Universal Robots URScript: swab_sampling.script

global swab_poses=make_list(0,0,6)
global pose_list_hor=make_list(0,0,420)
global pose_list_ver=make_list(0,0,420)
global cntd=False
global trgt_waypts=make_list(0,0,6)
global new_z=0
global first_pts=make_list(0,0,15)
global temp_pose_force=p[0,0,0,0,0,0]
global delta_rx=0
global new_dz=0
global server_msg=""
global delta_x=0
global delta_y=0


def connect2server():
	IP="192.168.12.139"
	port=3002
	while(cntd==False):
		cntd=socket_open(IP,port)
		if(cntd==True):
			textmsg("Connected to server")
		end
	end
	socket_send_string("SCAN_TARGET")
end


def get_hor_pose_from_server():

	IP="192.168.12.139"
	port=3002
	if(cntd==True):
		textmsg("Connected to server")
	end
	while(cntd==False):
		cntd=socket_open(IP,port)
		if(cntd==True):
			textmsg("Connected to server")
		end
		sleep(0.2)
	end
	socket_send_string("GET_POSE_HOR")
	idx=socket_read_ascii_float(1,timeout=-1)
	textmsg("Index from server=",idx[1])
	itn_i=0
	while(itn_i<idx[1]):
		msg=socket_read_ascii_float(6,timeout=-1)
		i=1
		while(i<7):
			swab_poses.append(msg[i])
			i=i+1
		end
		pose_list_hor.extend(swab_poses)
		swab_poses.clear()
		socket_send_string("OK")
		itn_i=itn_i+1
	end
	socket_read_line(timeout=-1)
	if(cntd==True):
		cntd=False
		socket_close()
	end
	#textmsg("server msg",swab_poses)
	textmsg("pose list",pose_list_hor)
end


def get_ver_pose_from_server():
	IP="192.168.12.139"
	port=3002
	if(cntd==True):
		textmsg("Connected to server")
	end
	while(cntd==False):
		cntd=socket_open(IP,port)
		if(cntd==True):
			textmsg("Connected to server")
		end
		sleep(0.2)
	end
	socket_send_string("GET_POSE_VER")
	idx=socket_read_ascii_float(1,timeout=-1)
	textmsg("Index from server=",idx[1])
	itn_i=0
	while(itn_i<idx[1]):
		msg=socket_read_ascii_float(6,timeout=-1)
		i=1
		while(i<7):
			swab_poses.append(msg[i])
			i=i+1
		end
		pose_list_ver.extend(swab_poses)
		swab_poses.clear()
		socket_send_string("OK")
		itn_i=itn_i+1
	end
	socket_read_line(timeout=-1)
	if(cntd==True):
		cntd=False
		socket_close()
	end
	#textmsg("server msg",swab_poses)
	textmsg("pose list",pose_list_ver)
end


def move_to_first_point(code):
	first_pts.clear()
	k=0
	i=1
	l=1
	blend_r=0
	while(i<3):
		j=1
		while(j<=6):
			k=l-1
			if(code==1):
				first_pts.append(pose_list_hor[k])
			elif(code==2):
				first_pts.append(pose_list_ver[k])
			end
			j=j+1
			l=l+1
		end
		i=i+1
	end
	movel(p[first_pts[0]-delta_y,first_pts[1]+delta_x,first_pts[2],first_pts[3],first_pts[4],first_pts[5]],a=0.5,v=0.05,r=blend_r)
	sleep(2)
	zero_ftsensor()
	sleep(2)
	tcp_f=get_tcp_force()
	textmsg("Force after zeroing:",tcp_f)
	ftmode=True
	while(ftmode==True):
		tcp_f=get_tcp_force()
		if tcp_f[2]<0.7:
			speedl([0,0,-0.001,0,0,0],0.05,t=0.5)
		else:
			stopl(3)
			new_p=get_actual_tcp_pose()
			new_z=new_p[2]-first_pts[2]
			ftmode=False
		end
		sleep(0.2)
	end
	movel(p[first_pts[6]-delta_y,first_pts[7]+delta_x,first_pts[8]+new_z,first_pts[9],first_pts[10],first_pts[11]],a=0.5,v=0.05,r=blend_r)
	curr_tcp=get_actual_tcp_pose()
	textmsg("Current TCP",curr_tcp)
	#tcp_str=to_string(curr_tcp)
	popup("Tcp change",blocking=True)
	#temp_pose_force=p[first_pts[0],first_pts[1],first_pts[2],first_pts[3],first_pts[4],first_pts[5]]
	temp_pt=first_pts[2]
	first_pts.clear()
	zero_ftsensor()
	sleep(2)
	tcp_f=get_tcp_force()
	textmsg("Force after zeroing:",tcp_f)
	ftmode=True
	#ftmode=False
	while(ftmode==True):
		tcp_f=get_tcp_force()
		textmsg("Force",tcp_f)
		if tcp_f[2]<2.5:
			speedl([0,0,-0.005,0,0,0],0.05,t=0.5)
		else:
			stopl(3)
			new_p=get_actual_tcp_pose()
			new_dz=new_p[2]-temp_pt
			ftmode=False
			textmsg("DZ=",new_dz)
		end
		sleep(0.2)
	end
	IP="192.168.12.139"
	port=3002
	if(cntd==True):
		textmsg("Connected to server")
	end
	while(cntd==False):
		cntd=socket_open(IP,port)
		if(cntd==True):
			textmsg("Connected to server")
		end
		sleep(0.2)
	end
	socket_send_string("POSE")
	socket_send_string(str_cat("",curr_tcp))
	if(cntd==True):
		cntd=False
		socket_close()
	end

end

def follow_swab_trajectory_hor():
	idx=pose_list_hor.length()
	textmsg("idx",idx)
	idx=idx/6
	k=0
	i=3
	l=13
	delta_z=0.035
	zero_ftsensor()
	sleep(1)
	#tcp_f=get_tcp_force()
	#textmsg("Force at tip:",tcp_f)
	force_mode(temp_pose_force,[0,0,1,0,0,0],[0,0,0.3,0,0,0],2,[0.005,0.005,0.05,0.01,0.01,0.01])
	while(i<=idx):
		j=1
		while(j<=6):
			k=l-1
			trgt_waypts.append(pose_list_hor[k])
			j=j+1
			l=l+1
		end
		if(i<3):
			delta_rx=0
			delta_z=0
			blend_r=0
		elif((i-1)%5==0):
			blend_r=0
			delta_z=0.043
			#delta_rx=0.104
			delta_rx=0.3
		else:
			blend_r=0.002
			delta_z=0.043
			#delta_rx=0.104
			delta_rx=0.3
		end
		if(i==1):
			delta_z=0.005
			trgt_waypts[2]=trgt_waypts[2]+delta_z
		movel(p[trgt_waypts[0],trgt_waypts[1],trgt_waypts[2],trgt_waypts[3],trgt_waypts[4],trgt_waypts[5]],a=0.5,v=0.05,r=blend_r)
			zero_ftsensor()
			sleep(1)
			ftmode=True
			while(ftmode==True):
				tcp_f=get_tcp_force()
				if tcp_f[2]<0.7:
					speedl([0,0,-0.001,0,0,0],0.5,t=0.5)
				else:
					stopl(3)
					new_p=get_actual_tcp_pose()
					new_z=new_p[2]-trgt_waypts[2]
					textmsg("Force at tip:",tcp_f)
					ftmode=False
				end
				sleep(0.2)
			end
		else:

			delta_z=0
			trgt_waypts[2]=trgt_waypts[2]+new_z+delta_z+new_dz
			trgt_waypts[3]=trgt_waypts[3]-delta_rx
		movel(p[trgt_waypts[0],trgt_waypts[1],trgt_waypts[2],trgt_waypts[3],trgt_waypts[4],trgt_waypts[5]],a=0.5,v=0.01,r=blend_r)
			tcp_f=get_tcp_force()
			#tcp_f=get_tcp_force_tool()
			textmsg("Force at tip:",tcp_f)
		end
		textmsg("Target Waypoints",trgt_waypts)
		trgt_waypts.clear()
		i=i+1
	end
	end_force_mode()
	pose_list_hor.clear()
end

def follow_swab_trajectory(code):
	dy=0.036
	pose_list_temp=make_list(0,0,420)
	if(code==1):
		pose_list_temp=pose_list_hor
		delta_x=0
		delta_y=0
	elif(code==2):
		pose_list_temp=pose_list_ver
	end
	idx=pose_list_temp.length()
	textmsg("idx",idx)
	idx=idx/6
	k=0
	i=3
	l=13

	zero_ftsensor()
	sleep(2)
	IP="192.168.12.139"
	port=3002
	if(cntd==True):
		textmsg("Connected to server")
	end
	while(cntd==False):
		cntd=socket_open(IP,port)
		if(cntd==True):
			textmsg("Connected to server")
		end
		sleep(0.2)
	end
	#force_mode(temp_pose_force,[0,0,1,0,0,0],[0,0,1,0,0,0],2,[0.001,0.001,0.01,0.01,0.01,0.01])
	while(i<=idx):
		socket_send_string("PLOT")
		j=1
		while(j<=6):
			k=l-1
			trgt_waypts.append(pose_list_temp[k])
			j=j+1
			l=l+1
		end
		if(i<3):
			delta_rx=0
			delta_z=0
			blend_r=0
		elif((i-1)%5==0):
			blend_r=0
			#delta_z=0.043
			#delta_rx=0.104
			delta_rx=0.3
		else:
			blend_r=0.002
			#delta_z=0.043
			#delta_rx=0.104
			delta_rx=0.3
		end
		delta_z=0
		if(i==3):
			temp=get_actual_tcp_pose()
			delta_y=temp[1]-trgt_waypts[1]
			delta_x=temp[0]-trgt_waypts[0]
		end
		#textmsg("delta Y:",delta_y)
		#textmsg("delta X:",delta_x)
		delta_x=0
		delta_y=0
		trgt_waypts[0]=trgt_waypts[0]+delta_x
		trgt_waypts[1]=trgt_waypts[1]+delta_y
		trgt_waypts[2]=trgt_waypts[2]+new_dz 		#new_z
		trgt_pose=pose_trans(p[trgt_waypts[0],trgt_waypts[1],trgt_waypts[2],trgt_waypts[3],trgt_waypts[4],trgt_waypts[5]],p[0,0,0,0,0,0])
		movel(trgt_pose,a=0.5,v=0.005,r=blend_r)
		tcp_f=get_tcp_force()
		#textmsg("Force at tip:",tcp_f)
		#textmsg("Target Waypoints",trgt_waypts)
		trgt_waypts.clear()
		i=i+1
	end
	#end_force_mode()
	socket_send_string("PLOT DONE")
	if(cntd==True):
		cntd=False
		socket_close()
	end
	#speedl([0,0,0.05,0,0,0],0.05,t=0.5)
	pose_list_temp.clear()
	if(code==2):
		delta_x=0
		delta_y=0
	end
end


def follow_swab_trajectory_ver():
	idx=pose_list_ver.length()
	textmsg("idx",idx)
	idx=idx/6
	k=0
	i=1
	l=1
	while(i<=idx):
		j=1
		while(j<=6):
			k=l-1
			trgt_waypts.append(pose_list_ver[k])
			j=j+1
			l=l+1
		end
		movel(p[trgt_waypts[0],trgt_waypts[1],trgt_waypts[2],trgt_waypts[3],trgt_waypts[4],trgt_waypts[5]],a=0.5,v=0.2)
		textmsg("Target Waypoints",trgt_waypts)
		trgt_waypts.clear()
		i=i+1
	end
	pose_list_ver.clear()
end


def wait_acknowledge():
	pose_list_hor.clear()
	pose_list_ver.clear()
	IP="192.168.12.139"
	port=3002
	if(cntd==True):
		textmsg("already Connected to server")
	end
	while(cntd==False):
		cntd=socket_open(IP,port)
		if(cntd==True):
			textmsg("Connected to server")
		end
		sleep(0.2)
	end
	serv_msg=socket_read_line(timeout=-1)
	textmsg("Server Message",serv_msg)

	if(cntd==True):
		cntd=False
		socket_close()
	end
	return serv_msg

end

def disconnectfromserver():
	delta_x=0
	delta_y=0
	socket_close()
end

def swab_break():
	curr_tcp=get_actual_tcp_pose()
	brk_pt=pose_add(curr_tcp,p[0,0,0.04,0,0,0])
	popup("tcp_changed to breaking point",blocking=True)
	movel(pose_trans(brk_pt,p[0,0,0,0,1.3,0]),a=0.5,v=0.005)
	#movel(p[brk_pt[0],brk_pt[1],brk_pt[02],brk_pt[3],brk_pt[4]+1.57,brk_pt[5]],a=0.5,v=0.005)
end

#Helper Function

def get_tcp_force_tool():
	force_torque= get_tcp_force()
	force_B=p[force_torque[0],force_torque[1],force_torque[2],0,0,0]
	torque_B=p[force_torque[3],force_torque[4],force_torque[5],0,0,0]
	tcp=temp_pose_force
	rotation_BT=p[0,0,0,tcp[3],tcp[4],tcp[5]]
	force_T= pose_trans(pose_inv(rotation_BT),force_B)
	torque_T=pose_trans(pose_inv(rotation_BT),torque_B)
	force_torque_T=p[force_T[0],force_T[1],force_T[2],torque_T[0],torque_T[1],torque_T[2]]
	return force_torque_T
end
